Fanuc KAREL source: ka00175.KL

PROGRAM KA00175
%STACKSIZE=65535
%PRIORITY=65535
%NOLOCKGROUP
VAR
SRC : ARRAY[4] OF STRING[20]
DST : ARRAY[4] OF STRING[20]
BEGIN
-- UNRESOLVED_PC line 7 opcodes [22 22 1E] marker_code=0
END KA00175
